FUNCTION_BLOCK SENSOR_ADCPI
  {SET_ATTRIBUTE(OpcUa, DEVICE.SENSOR)}
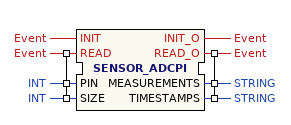
  EVENT_INPUT
    INIT;
    READ WITH PIN, SIZE;
  END_EVENT
  EVENT_OUTPUT
    INIT_O;
    READ_O WITH MEASUREMENTS, TIMESTAMPS;
  END_EVENT
  VAR_INPUT
    PIN : INT; {SET_ATTRIBUTE(OpcUa, Variable)}
    SIZE : INT; {SET_ATTRIBUTE(OpcUa, Variable)}
  END_VAR
  VAR_OUTPUT
    MEASUREMENTS : STRING; {SET_ATTRIBUTE(OpcUa, Variable)}
    TIMESTAMPS : STRING; {SET_ATTRIBUTE(OpcUa, Variable)}
  END_VAR
END_FUNCTION_BLOCK
